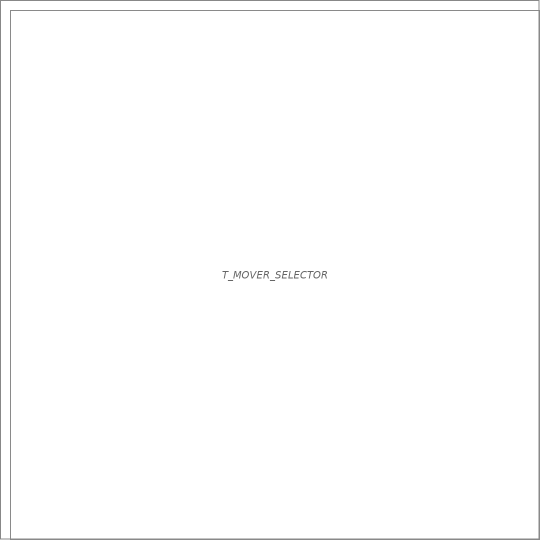
VISUALIZATION SELECTOR_VISU  // 540x540
    Frame (10,10 530x530)
        shows T_MOVER_SELECTOR(Control := GVL_XTS.MoverSelectorCtrl, State := GVL_XTS.MoverSelectorState, sState := GVL_APPLICATION.VisuPoolData.sSelectorState, sResult := GVL_APPLICATION.VisuPoolData.sSelectorResult)
END_VISUALIZATION

(* stored: Version 1.1.0.1
   Visu SELECTOR_VISU: Id {9ad0cb5c-0a74-4dff-85d6-b6a2f3f3400f} *)
